// Mitsubishi GX Works2 project: Main Program   PLC: FX3U/FX3UC

PROGRAM MAIN
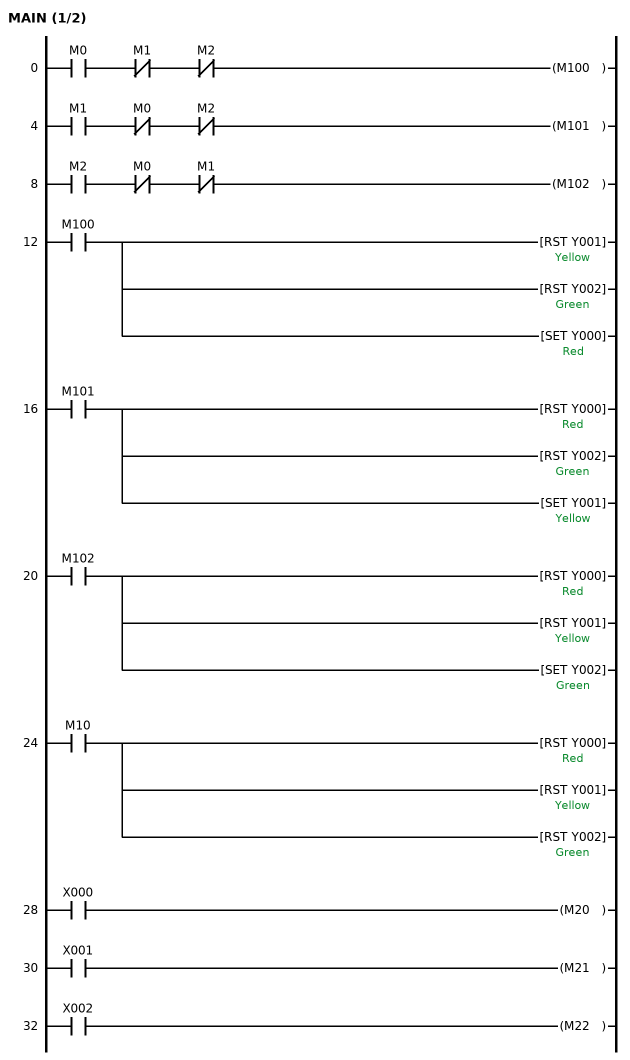
0     LD      M0
      ANI     M1
      ANI     M2
      OUT     M100
4     LD      M1
      ANI     M0
      ANI     M2
      OUT     M101
8     LD      M2
      ANI     M0
      ANI     M1
      OUT     M102
12    LD      M100
      RST     Y001  ; Yellow
      RST     Y002  ; Green
      SET     Y000  ; Red
16    LD      M101
      RST     Y000  ; Red
      RST     Y002  ; Green
      SET     Y001  ; Yellow
20    LD      M102
      RST     Y000  ; Red
      RST     Y001  ; Yellow
      SET     Y002  ; Green
24    LD      M10
      RST     Y000  ; Red
      RST     Y001  ; Yellow
      RST     Y002  ; Green
28    LD      X000
      OUT     M20
30    LD      X001
      OUT     M21
32    LD      X002
      OUT     M22
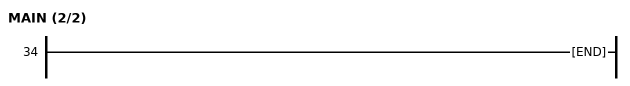
34    END
END_PROGRAM
